(* IEC 61131-3 sources: STEPROBOT/docs/welder_r6_4/source_reference, 3 files *)

(* ---- CommPoll.declaration.original.st ---- *)
(* ================================================================ *)
(* InoProShop 创建方式:                                              *)
(*   右键 Application → 添加对象 → 程序(POU)                        *)
(*   名称: CommPoll, 语言: ST, 类型: PROGRAM                        *)
(*   任务分配: MainTask (1ms周期)                                    *)
(*   说明: 焊机EtherCAT I/O 周期打包/解析                            *)
(*   依赖GVL: GVL_Welder, GVL_CNC                                  *)
(* ================================================================ *)
(*
 * 职责划分:
 *   CNC_Main.st  → 仅设置布尔标志 (g_wWeldOn, g_wRobotReady等)
 *   CommPoll.st  → 每周期: D300拆位→独立BOOL→组装g_byWeldOut
 *                    独立BOOL→组装D308+解析g_byWeldIn
 *
 * 字节映射依据: 奥太EtherCAT通讯协议 2024.7.1
 * PLC数组下标 = 协议字节号 (0-based)
 * ================================================================ *)

PROGRAM CommPoll
VAR
    nTempU16 : UINT;
    nTempI16 : INT;
    byTemp   : BYTE;
    wCtrlPacked : UINT;
    wPrevCtrlPacked : UINT := 16#FFFF;
    bBootInit : BOOL := TRUE;
    rPrevWireAuto : REAL;
    lrPrevWireRun : LREAL;
    bWireParamInit : BOOL := TRUE;
END_VAR

(* ---- CommPoll.implementation.original.st ---- *)
(* Canonical wire parameters: reject NaN/infinity/negative values without
   converting them to integer timer values. No command/enable is generated. *)
IF NOT ((g_rWireStartDelay >= 0.0) AND (g_rWireStartDelay <= 60.0)) THEN
    g_rWireStartDelay := 0.0;
END_IF;
IF NOT ((g_rWireStopDelay >= 0.0) AND (g_rWireStopDelay <= 60.0)) THEN
    g_rWireStopDelay := 0.0;
END_IF;
IF NOT ((g_rWireJogSpeed >= 0.0) AND (g_rWireJogSpeed <= 1000.0)) THEN
    g_rWireJogSpeed := 0.0;
END_IF;
IF NOT ((g_rWireAutoSpeed >= 0.0) AND (g_rWireAutoSpeed <= 1000.0)) THEN
    g_rWireAutoSpeed := 0.0;
END_IF;
IF NOT ((g_fWireFeedSpeed >= 0.0) AND (g_fWireFeedSpeed <= 1000.0)) THEN
    g_fWireFeedSpeed := 0.0;
END_IF;
IF bWireParamInit THEN
    (* Preserve the existing 64-bit setting across restart. *)
    g_rWireAutoSpeed := LREAL_TO_REAL(g_fWireFeedSpeed);
    bWireParamInit := FALSE;
ELSIF g_fWireFeedSpeed <> lrPrevWireRun THEN
    g_rWireAutoSpeed := LREAL_TO_REAL(g_fWireFeedSpeed);
ELSIF g_rWireAutoSpeed <> rPrevWireAuto THEN
    g_fWireFeedSpeed := REAL_TO_LREAL(g_rWireAutoSpeed);
END_IF;
rPrevWireAuto := g_rWireAutoSpeed;
lrPrevWireRun := g_fWireFeedSpeed;
g_dwModbusSignature := 16#4D573031;
g_wModbusMapVersion := 1;
g_dwModbusCycle := g_dwModbusCycle + UDINT#1;
g_wModbusProbeEcho := g_wModbusProbe XOR UINT#16#A55A;

IF bBootInit THEN
    g_wWeldCtrlWord := 0;
    g_wWeldOn := FALSE;
    g_wRobotReady := FALSE;
    g_wGasCheck := FALSE;
    g_bHotWireEnable := FALSE;
    g_bHotWireACMode := FALSE;
    g_bHighFreqDisable := FALSE;
    g_bGunCoolMode := FALSE;
    wPrevCtrlPacked := 0;
    bBootInit := FALSE;
END_IF;

(* ================================================================ *)
(* D300 <-> 独立BOOL 双向合并                                         *)
(* 1. 从独立BOOL打包到临时变量                                        *)
(* 2. 若D300与上次打包值不同(PC写了D300), 则拆位D300→BOOL             *)
(* 3. 再从BOOL打包→D300 (PLC改BOOL也能反映到D300)                     *)
(* ================================================================ *)

wCtrlPacked := 0;
IF g_wWeldOn         THEN wCtrlPacked := wCtrlPacked OR 16#0001; END_IF;
IF g_wRobotReady     THEN wCtrlPacked := wCtrlPacked OR 16#0002; END_IF;
IF g_wGasCheck       THEN wCtrlPacked := wCtrlPacked OR 16#0004; END_IF;
IF g_bHotWireEnable  THEN wCtrlPacked := wCtrlPacked OR 16#0008; END_IF;
IF g_bHotWireACMode  THEN wCtrlPacked := wCtrlPacked OR 16#0010; END_IF;
IF g_bHighFreqDisable THEN wCtrlPacked := wCtrlPacked OR 16#0080; END_IF;
IF g_bGunCoolMode    THEN wCtrlPacked := wCtrlPacked OR 16#0100; END_IF;

IF g_wWeldCtrlWord <> wPrevCtrlPacked THEN
    g_wWeldOn         := (g_wWeldCtrlWord AND 16#0001) <> 0;
    g_wRobotReady     := (g_wWeldCtrlWord AND 16#0002) <> 0;
    g_wGasCheck       := (g_wWeldCtrlWord AND 16#0004) <> 0;
    g_bHotWireEnable  := (g_wWeldCtrlWord AND 16#0008) <> 0;
    g_bHotWireACMode  := (g_wWeldCtrlWord AND 16#0010) <> 0;
    g_bHighFreqDisable := (g_wWeldCtrlWord AND 16#0080) <> 0;
    g_bGunCoolMode    := (g_wWeldCtrlWord AND 16#0100) <> 0;
    wCtrlPacked := g_wWeldCtrlWord;
END_IF;

g_wWeldCtrlWord := wCtrlPacked;
wPrevCtrlPacked := wCtrlPacked;

(* ================================================================ *)
(* 焊机输出 (协议: 焊机的输入数据区, PLC写→焊机读)                    *)
(* g_byWeldOut[0..31] → EtherCAT输出 → 焊机                        *)
(* ================================================================ *)

(* ===== 协议 Byte 0: 控制位 ===== *)
(* bit0(1):  开始焊接 1=起弧 0=停弧                                  *)
(* bit1(2):  机器人准备好 高有效                                      *)
(* bit2(3):  检气 高有效                                              *)
(* bit3-4:   焊机操作模式 00=两步 01=四步 10=反复                     *)
(* bit5-7:   焊机工作模式 000=直流恒流 001=直流脉冲 010=交流恒流       *)
(*           011=交流脉冲 100=直流手弧焊                               *)
byTemp := 0;
IF g_wWeldOn THEN byTemp := byTemp OR 16#01; END_IF;
IF g_wRobotReady THEN byTemp := byTemp OR 16#02; END_IF;
IF g_wGasCheck THEN byTemp := byTemp OR 16#04; END_IF;
nTempU16 := LIMIT(UINT#0, g_wWeldOperMode, UINT#2);
byTemp := byTemp OR SHL(UINT_TO_BYTE(nTempU16), 3);
nTempU16 := LIMIT(UINT#0, g_wWeldWorkMode, UINT#4);
byTemp := byTemp OR SHL(UINT_TO_BYTE(nTempU16), 5);
g_byWeldOut[0] := byTemp;

(* ===== 协议 Byte 1: 辅助控制位 ===== *)
(* bit0(9):  热丝电源使能 1=ON 0=OFF                                  *)
(* bit1(10): 热丝工作模式 0=DC 1=AC                                   *)
(* bit2(11): 备用                                                     *)
(* bit3(12): 点动送丝 (已移除, 送丝通过轴控制) *)
(* bit4(13): 点动抽丝 (已移除, 送丝通过轴控制) *)
(* bit5(14): 备用                                                     *)
(* bit6(15): 高频有无 0=高频 1=提升                                   *)
(* bit7(16): 焊枪模式 0=水冷 1=气冷                                   *)
byTemp := 0;
IF g_bHotWireEnable THEN byTemp := byTemp OR 16#01; END_IF;
IF g_bHotWireACMode THEN byTemp := byTemp OR 16#02; END_IF;
IF g_bHighFreqDisable THEN byTemp := byTemp OR 16#40; END_IF;
IF g_bGunCoolMode THEN byTemp := byTemp OR 16#80; END_IF;
g_byWeldOut[1] := byTemp;

(* ===== 协议 Byte 2: 热丝频率 ===== *)
(* 范围: 20-100 对应20~100Hz (1字节) *)
g_byWeldOut[2] := UINT_TO_BYTE(LIMIT(UINT#20, g_wHotWireFreq, UINT#100));

(* ===== 协议 Byte 3: 热丝电流给定 ===== *)
(* 范围: 0-200 对应0~200A (1字节) *)
g_byWeldOut[3] := UINT_TO_BYTE(LIMIT(UINT#0, g_wHotWireCurrent, UINT#200));

(* ===== 协议 Byte 4-5: 给定电流 (2字节小端, 低字节在前) ===== *)
(* 范围: 40-4000 对应4.0~400.0A *)
nTempU16 := REAL_TO_UINT(LIMIT(4.0, g_wWeldCurrent, 400.0)*10.0);

g_byWeldOut[4] := UINT_TO_BYTE(UINT_TO_USINT(nTempU16 MOD 256));
g_byWeldOut[5] := UINT_TO_BYTE(UINT_TO_USINT(nTempU16 / 256));

(* ===== 协议 Byte 6: 送丝速度 (已移除, 送丝通过轴控制, 写0) ===== *)
g_byWeldOut[6] := 0;

(* ===== 协议 Byte 7: 起弧延迟送丝时间 (已移除, 写0) ===== *)
g_byWeldOut[7] := 0;

(* ===== 协议 Byte 8: 熄弧滞后送丝时间 (已移除, 写0) ===== *)
g_byWeldOut[8] := 0;

(* ===== 协议 Byte 9: 熄弧回抽丝长度 (已移除, 写0) ===== *)
g_byWeldOut[9] := 0;

(* ===== 协议 Byte 10: 点动送丝速度 (已移除, 送丝通过轴控制, 写0) ===== *)
g_byWeldOut[10] := 0;

(* ===== 协议 Byte 11: 通讯异常标志 (控制器填充) ===== *)
g_byWeldOut[11] := g_wCommErrorFlag;

(* ===== 协议 Byte 12: 慢送丝速度 (已移除, 送丝通过轴控制, 写0) ===== *)
g_byWeldOut[12] := 0;

(* ===== 协议 Byte 13-14: 前气时间 (2字节小端, 低字节在前) ===== *)
(* 范围: 1-999 对应0.01~9.99s *)
nTempU16 := REAL_TO_UINT(LIMIT(0.01, g_wFrontGasTime, 9.99)*100.0);
g_byWeldOut[13] := UINT_TO_BYTE(UINT_TO_USINT(nTempU16 MOD 256));
g_byWeldOut[14] := UINT_TO_BYTE(UINT_TO_USINT(nTempU16 / 256));

(* ===== 协议 Byte 15-16: 延气时间 (2字节小端, 低字节在前) ===== *)
(* 范围: 1-600 对应0.1~60.0s *)
nTempU16 := REAL_TO_UINT(LIMIT(0.1, g_wTailGasTime, 60.0)*10.0);
g_byWeldOut[15] := UINT_TO_BYTE(UINT_TO_USINT(nTempU16 MOD 256));
g_byWeldOut[16] := UINT_TO_BYTE(UINT_TO_USINT(nTempU16 / 256));

(* ===== 协议 Byte 17: 爬升时间 ===== *)
(* 范围: 1-100 对应0.1~10.0s (1字节) *)
g_byWeldOut[17] := UINT_TO_BYTE(REAL_TO_UINT(LIMIT(0.1, g_wRampUpTime, 10.0)*10.0));

(* ===== 协议 Byte 18: 衰减时间 ===== *)
(* 范围: 1-150 对应0.1~15.0s (1字节) *)
g_byWeldOut[18] := UINT_TO_BYTE(REAL_TO_UINT(LIMIT(0.1, g_wRampDownTime, 15.0)*10.0));

(* ===== 协议 Byte 19: 脉冲频率 ===== *)
(* 范围: 2-200 对应0.2~20.0Hz (1字节) *)
g_byWeldOut[19] := UINT_TO_BYTE(REAL_TO_UINT(LIMIT(0.2, g_wPulseFreq, 20.0)*10.0));

(* ===== 协议 Byte 20-22: 占空比 + 峰值电流 (交叉编排) ===== *)
(* 占空比: Byte20=低字节, Byte22 bit4-7=高字节低4位 (范围1-999, 12位) *)
(* 峰值电流: Byte21=低字节, Byte22 bit0-3=高字节低4位 (范围50-4000, 12位) *)
(* 占空比 = [Byte22 bit7:4][Byte20] *)
(* 峰值电流 = [Byte22 bit3:0][Byte21] *)
nTempU16 := REAL_TO_UINT(LIMIT(0.1, g_wDutyCycle, 99.9)*10.0);
g_byWeldOut[20] := UINT_TO_BYTE(UINT_TO_USINT(nTempU16 MOD 256));
g_byWeldOut[21] := UINT_TO_BYTE(UINT_TO_USINT(REAL_TO_UINT(LIMIT(5.0, g_wPeakCurrent, 400.0)*10.0) MOD 256));
byTemp := 0;
byTemp := byTemp OR SHL(UINT_TO_BYTE(UINT_TO_USINT(nTempU16 / 256)) AND 16#0F, 4);
byTemp := byTemp OR (UINT_TO_BYTE(UINT_TO_USINT(REAL_TO_UINT(LIMIT(5.0, g_wPeakCurrent, 400.0)*10.0) / 256)) AND 16#0F);
g_byWeldOut[22] := byTemp;

(* ===== 协议 Byte 23-24: 基值电流 (2字节小端, 低字节在前) ===== *)
(* 范围: 50-4000 对应5.0~400.0A *)
nTempU16 := REAL_TO_UINT(LIMIT(5.0, g_wBaseCurrent, 400.0)*10.0);
g_byWeldOut[23] := UINT_TO_BYTE(UINT_TO_USINT(nTempU16 MOD 256));
g_byWeldOut[24] := UINT_TO_BYTE(UINT_TO_USINT(nTempU16 / 256));

(* ===== 协议 Byte 25-26: 起弧电流 (2字节小端, 低字节在前) ===== *)
(* 范围: 50-4000 对应5.0~400.0A *)
nTempU16 := REAL_TO_UINT(LIMIT(5.0, g_wArcStartCurrent, 400.0)*10.0);
g_byWeldOut[25] := UINT_TO_BYTE(UINT_TO_USINT(nTempU16 MOD 256));
g_byWeldOut[26] := UINT_TO_BYTE(UINT_TO_USINT(nTempU16 / 256));

(* ===== 协议 Byte 27-28: 收弧电流 (2字节小端, 低字节在前) ===== *)
(* 范围: 50-4000 对应5.0~400.0A *)
nTempU16 := REAL_TO_UINT(LIMIT(5.0, g_wArcEndCurrent, 400.0)*10.0);
g_byWeldOut[27] := UINT_TO_BYTE(UINT_TO_USINT(nTempU16 MOD 256));
g_byWeldOut[28] := UINT_TO_BYTE(UINT_TO_USINT(nTempU16 / 256));

(* ===== 协议 Byte 29: 交流频率 ===== *)
(* 范围: 40-250 对应40-250Hz (1字节) *)
g_byWeldOut[29] := UINT_TO_BYTE(LIMIT(UINT#40, g_wACFreq, UINT#250));

(* ===== 协议 Byte 30: 清理比例 ===== *)
(* 范围: 90-180 对应40~-50 (1字节) *)
nTempI16 := 130 - UINT_TO_INT(LIMIT(UINT#90, g_wCleanRatio, UINT#180));
g_byWeldOut[30] := INT_TO_BYTE(nTempI16);

(* ===== 协议 Byte 31: 交流偏置 ===== *)
(* 范围: 90-180 对应40~-50 (1字节) *)
nTempI16 := 130 - UINT_TO_INT(LIMIT(UINT#90, g_wACBias, UINT#180));
g_byWeldOut[31] := INT_TO_BYTE(nTempI16);

(* ================================================================ *)
(* 焊机输入 (协议: 焊机输出数据区, 焊机写→PLC读)                      *)
(* g_byWeldIn[0..31] ← EtherCAT输入 ← 焊机                          *)
(* ================================================================ *)

(* ===== 协议输入 Byte 0: 状态位 ===== *)
(* bit0: 引弧成功 高有效                                              *)
(* bit1: 焊机准备好 高有效                                            *)
(* bit2: 预留                                                         *)
(* bit3: 电流有无 高有效                                              *)
(* EtherCAT 输入映射别名 → 协议数组。保持原有 Byte 0..31 定义。 *)
g_byWeldIn[0] := g_byWeldInMap01;
g_byWeldIn[1] := g_byWeldInMap02;
g_byWeldIn[2] := g_byWeldInMap03;
g_byWeldIn[3] := g_byWeldInMap04;
g_byWeldIn[4] := g_byWeldInMap05;
g_byWeldIn[5] := g_byWeldInMap06;
g_byWeldIn[6] := g_byWeldInMap07;
g_byWeldIn[7] := g_byWeldInMap08;
g_byWeldIn[8] := g_byWeldInMap09;
g_byWeldIn[9] := g_byWeldInMap10;
g_byWeldIn[10] := g_byWeldInMap11;
g_byWeldIn[11] := g_byWeldInMap12;
g_byWeldIn[12] := g_byWeldInMap13;
g_byWeldIn[13] := g_byWeldInMap14;
g_byWeldIn[14] := g_byWeldInMap15;
g_byWeldIn[15] := g_byWeldInMap16;
g_byWeldIn[16] := g_byWeldInMap17;
g_byWeldIn[17] := g_byWeldInMap18;
g_byWeldIn[18] := g_byWeldInMap19;
g_byWeldIn[19] := g_byWeldInMap20;
g_byWeldIn[20] := g_byWeldInMap21;
g_byWeldIn[21] := g_byWeldInMap22;
g_byWeldIn[22] := g_byWeldInMap23;
g_byWeldIn[23] := g_byWeldInMap24;
g_byWeldIn[24] := g_byWeldInMap25;
g_byWeldIn[25] := g_byWeldInMap26;
g_byWeldIn[26] := g_byWeldInMap27;
g_byWeldIn[27] := g_byWeldInMap28;
g_byWeldIn[28] := g_byWeldInMap29;
g_byWeldIn[29] := g_byWeldInMap30;
g_byWeldIn[30] := g_byWeldInMap31;
g_byWeldIn[31] := g_byWeldInMap32;

g_bWeldArcOK      := (g_byWeldIn[0] AND 16#01) <> 0;
g_bWeldReady      := (g_byWeldIn[0] AND 16#02) <> 0;
g_bWeldHasCurrent     := (g_byWeldIn[0] AND 16#08) <> 0;

(* ===== 协议输入 Byte 1: 报警位 ===== *)
(* bit0: 预留                                                         *)
(* bit1: 焊枪开关异常 高有效                                          *)
(* bit2: 焊机热保护 高有效                                            *)
(* bit3: 缺水保护 高有效                                              *)
(* bit4: 热丝电源热保护 高有效                                        *)
(* bit5: 热丝电源通讯保护 高有效 (控制器填充)                          *)
g_bGunSwitchFault    := (g_byWeldIn[1] AND 16#02) <> 0;
g_bWeldThermalProtect := (g_byWeldIn[1] AND 16#04) <> 0;
g_bWaterProtect   := (g_byWeldIn[1] AND 16#08) <> 0;
g_bWirePSThermal  := (g_byWeldIn[1] AND 16#10) <> 0;
g_bWirePSCommFault:= (g_byWeldIn[1] AND 16#20) <> 0;

(* ===== 报警组合 ===== *)
g_bWeldFault := g_bWeldThermalProtect
              OR g_bGunSwitchFault
              OR g_bWaterProtect
              OR g_bWirePSThermal
              OR g_bWirePSCommFault;

IF g_bWeldFault THEN
    g_rWeldFaultCode := BYTE_TO_UINT(g_byWeldIn[1]);
ELSE
    g_rWeldFaultCode := 0;
END_IF;

IF NOT g_bWeldReady OR g_bWeldFault THEN
    g_wWeldOn := FALSE;
    g_wWeldCtrlWord := g_wWeldCtrlWord AND 16#FFFE;
    wPrevCtrlPacked := wPrevCtrlPacked AND 16#FFFE;
    g_byWeldOut[0] := g_byWeldOut[0] AND 16#FE;
END_IF;

(* ===== EtherCAT 输出映射别名同步 ===== *)
(* 放在未就绪/故障联锁之后，确保停弧命令在本周期立即写入PDO。 *)
g_byWeldOutMap01 := g_byWeldOut[0];
g_byWeldOutMap02 := g_byWeldOut[1];
g_byWeldOutMap03 := g_byWeldOut[2];
g_byWeldOutMap04 := g_byWeldOut[3];
g_byWeldOutMap05 := g_byWeldOut[4];
g_byWeldOutMap06 := g_byWeldOut[5];
g_byWeldOutMap07 := g_byWeldOut[6];
g_byWeldOutMap08 := g_byWeldOut[7];
g_byWeldOutMap09 := g_byWeldOut[8];
g_byWeldOutMap10 := g_byWeldOut[9];
g_byWeldOutMap11 := g_byWeldOut[10];
g_byWeldOutMap12 := g_byWeldOut[11];
g_byWeldOutMap13 := g_byWeldOut[12];
g_byWeldOutMap14 := g_byWeldOut[13];
g_byWeldOutMap15 := g_byWeldOut[14];
g_byWeldOutMap16 := g_byWeldOut[15];
g_byWeldOutMap17 := g_byWeldOut[16];
g_byWeldOutMap18 := g_byWeldOut[17];
g_byWeldOutMap19 := g_byWeldOut[18];
g_byWeldOutMap20 := g_byWeldOut[19];
g_byWeldOutMap21 := g_byWeldOut[20];
g_byWeldOutMap22 := g_byWeldOut[21];
g_byWeldOutMap23 := g_byWeldOut[22];
g_byWeldOutMap24 := g_byWeldOut[23];
g_byWeldOutMap25 := g_byWeldOut[24];
g_byWeldOutMap26 := g_byWeldOut[25];
g_byWeldOutMap27 := g_byWeldOut[26];
g_byWeldOutMap28 := g_byWeldOut[27];
g_byWeldOutMap29 := g_byWeldOut[28];
g_byWeldOutMap30 := g_byWeldOut[29];
g_byWeldOutMap31 := g_byWeldOut[30];
g_byWeldOutMap32 := g_byWeldOut[31];

(* ===== 协议输入 Byte 4-5: 实际焊接电压 (2字节小端, 0.1V分辨率) ===== *)
(* 范围: 0-1000 对应0~100.0V *)
nTempU16 := BYTE_TO_UINT(g_byWeldIn[4]) + BYTE_TO_UINT(g_byWeldIn[5]) * 256;
g_rWeldVoltageAct := UINT_TO_REAL(nTempU16) * 0.1;

(* ===== 协议输入 Byte 6-7: 实际焊接电流 (2字节小端, 0.1A分辨率) ===== *)
(* 范围: 0~400 对应0~400A *)
nTempU16 := BYTE_TO_UINT(g_byWeldIn[6]) + BYTE_TO_UINT(g_byWeldIn[7]) * 256;
g_rWeldCurrentAct := UINT_TO_REAL(nTempU16) * 0.1;

(* ===== 协议输入 Byte 8-9: 实际热丝焊接电流 (2字节小端, 10A分辨率) ===== *)
(* 范围: 0~20 对应0~200A *)
nTempU16 := BYTE_TO_UINT(g_byWeldIn[8]) + BYTE_TO_UINT(g_byWeldIn[9]) * 256;
g_rHotWireCurrentAct := UINT_TO_REAL(nTempU16) * 10.0;

(* ===== 协议输入 Byte 10-11: 送丝速度反馈 (已移除, 送丝通过轴控制) ===== *)

(* ===== 组装输入状态字 (PC通过D500读取) ===== *)
g_wWeldInStatus := 0;
IF g_bWeldArcOK      THEN g_wWeldInStatus := g_wWeldInStatus OR 16#0001; END_IF;
IF g_bWeldReady      THEN g_wWeldInStatus := g_wWeldInStatus OR 16#0002; END_IF;
IF g_bGunSwitchFault THEN g_wWeldInStatus := g_wWeldInStatus OR 16#0004; END_IF;
IF g_bWeldThermalProtect THEN g_wWeldInStatus := g_wWeldInStatus OR 16#0008; END_IF;
IF g_bWaterProtect   THEN g_wWeldInStatus := g_wWeldInStatus OR 16#0010; END_IF;
IF g_bWirePSThermal  THEN g_wWeldInStatus := g_wWeldInStatus OR 16#0020; END_IF;
IF g_bWirePSCommFault THEN g_wWeldInStatus := g_wWeldInStatus OR 16#0040; END_IF;
IF g_bWeldFault      THEN g_wWeldInStatus := g_wWeldInStatus OR 16#0080; END_IF;
IF g_bWeldHasCurrent     THEN g_wWeldInStatus := g_wWeldInStatus OR 16#0100; END_IF;

(* ================================================================ *)
(* D308 独立BOOL → 打包字 (PLC内部 → PC读D308)                         *)
(* CommPoll每周期从独立BOOL组装到g_wWeldStatusWord供PC读取             *)
(* ================================================================ *)
g_wWeldStatusWord := 0;
IF g_bWeldArcOK      THEN g_wWeldStatusWord := g_wWeldStatusWord OR 16#0001; END_IF;
IF g_bWeldReady      THEN g_wWeldStatusWord := g_wWeldStatusWord OR 16#0002; END_IF;
IF g_bWeldHasCurrent     THEN g_wWeldStatusWord := g_wWeldStatusWord OR 16#0004; END_IF;
IF g_bGunSwitchFault THEN g_wWeldStatusWord := g_wWeldStatusWord OR 16#0008; END_IF;
IF g_bWeldThermalProtect THEN g_wWeldStatusWord := g_wWeldStatusWord OR 16#0010; END_IF;
IF g_bWaterProtect   THEN g_wWeldStatusWord := g_wWeldStatusWord OR 16#0020; END_IF;
IF g_bWirePSThermal  THEN g_wWeldStatusWord := g_wWeldStatusWord OR 16#0040; END_IF;
IF g_bWirePSCommFault THEN g_wWeldStatusWord := g_wWeldStatusWord OR 16#0080; END_IF;
IF g_bWeldFault      THEN g_wWeldStatusWord := g_wWeldStatusWord OR 16#0100; END_IF;

(* ================================================================ *)
(* 激光距离读取和转换                                                *)
(* 从%IW50读取激光距离原始INT值, 转换为实际距离并存入寄存器            *)
(* 转换公式: 实际距离 = 原始值 / 100 + 50                             *)
(* D522 = g_rLaserDistance (REAL, PC可通过Modbus读取)                   *)
(* ================================================================ *)
g_rLaserDistance := INT_TO_REAL(g_iLaserDistanceRaw) / 100.0 + 50.0;

(* ---- GVL_Welders.original.st ---- *)
(* EtherCAT -9 welder: 32-byte RxPDO/TxPDO use symbolic channel mappings; no fixed IEC addresses. *)
(* ================================================================ *)
(* InoProShop 创建方式:                                              *)
(*   右键 Application → 添加对象 → 全局变量表(GVL)                    *)
(*   名称: GVL_Welders                                               *)
(*   说明: 奥太焊机 EtherCAT 通讯接口全局变量                         *)
(*   依赖: 无                                                        *)
(*   修订: 布尔变量使用独立%MW地址 (D300控制=%MW101~109)               *)
(*         (D308状态=%MW111~119), InoProShop不支持BOOL位打包         *)
(*         新增 %MW300/%MW308 作为Modbus从站打包字映射 (方案C)         *)
(* ================================================================ *)
(*
 * EtherCAT通讯协议 (奥太 2024.7.1)
 *
 * EtherCAT输出 (PLC→焊机): g_byWeldOut[0..31] → 地址-9焊机RxPDO (32字节)
 *   协议字节0~31 = PLC数组下标0~31 (一一对应)
 *
 * EtherCAT输入 (焊机→PLC): g_byWeldIn[0..31] ← 地址-9焊机TxPDO (32字节)
 *   协议字节0~31 = PLC数组下标0~31 (一一对应)
 *
 * 数据流:
 *   PC(Modbus写D300) → g_wWeldCtrlWord (打包字)
 *       → CommPoll.st拆位 → g_wWeldOn等独立BOOL
 *       → CommPoll.st组装 → g_byWeldOut → EtherCAT → 焊机
 *   焊机 → EtherCAT → g_byWeldIn
 *       → CommPoll.st解析 → g_bWeldArcOK等独立BOOL
 *       → CommPoll.st组装 → g_wWeldStatusWord → PC(Modbus读D308)
 *
 * Modbus寄存器布局:
 *   D300 (%MW300): 焊机控制输出标志位 (16位打包字, CommPoll双向映射)
 *     独立BOOL: g_wWeldOn(%MW101) ~ g_bGunCoolMode(%MW109)
 *   D302      : 焊机操作模式 (UINT)
 *   D304      : 焊机工作模式 (UINT)
 *   D306      : 通讯异常标志 (BYTE, 控制器填充)
 *   D308 (%MW308): 焊机输入状态标志位 (16位打包字, CommPoll组装)
 *     独立BOOL: g_bWeldArcOK(%MW111) ~ g_bWeldFault(%MW119)
 *   D400-D444 : 焊接参数 (各参数见注释)
 *   D500      : 焊机输入状态字 (16位打包, CommPoll从独立BOOL组装)
 *   D502-D518 : 焊机输入反馈值
 *
 * 注意: Modbus从站配置需包含 D300-D306 和 D308 映射范围
 *       D300=%MW300, D308=%MW308 均为打包字, PC按位操作
 * ================================================================ *)

(* ================================================================= *)
(* 焊机控制输出标志位 → 协议 Byte 0 / Byte 1 位域                     *)
(* Modbus: D300 (%MW300, 16位), bit0~8 对应9个布尔量                  *)
(* ================================================================= *)

(*
 * 协议 Byte 0 位域:
 *   bit0(1):  开始焊接       1=起弧 0=停弧 [危险, 高有效]
 *   bit1(2):  机器人准备好   上位机接收到焊机数据, 通讯正常, 高有效
 *   bit2(3):  检气           高有效
 *   bit3-4:   焊机操作模式   00=两步 01=四步 10=反复
 *   bit5-7:   焊机工作模式   000=直流恒流 001=直流脉冲 010=交流恒流
 *             011=交流脉冲 100=直流手弧焊
 *
 * 协议 Byte 1 位域:
 *   bit0(9):  热丝电源使能   1=ON 0=OFF
 *   bit1(10): 热丝工作模式   0=DC 1=AC
 *   bit2(11): 备用
 *   bit3(12): 点动送丝       高有效, 丝检时使用, 电平信号
 *   bit4(13): 点动抽丝       高有效, 丝检时使用, 电平信号
 *   bit5(14): 备用
 *   bit6(15): 高频有无       0=高频 1=提升
 *   bit7(16): 焊枪模式       0=水冷 1=气冷
 *)

(* --- 协议 Byte 11: 通讯异常标志 (控制器填充) --- *)
(*
 * 协议 Byte 11 位域:
 *   bit0(89):  机器人→CAN控制器通信异常 (控制器填充, 焊机显示E84)
 *             注: 500ms内无机器人准备好信号将触发此异常
 *   bit1-3:    预留
 *   bit4(93):  焊机→CAN控制器通信异常 (控制器填充, 焊机显示E85)
 *   bit5-7:    预留
 *)

(* ================================================================= *)
(* 焊接参数 Modbus 接收 (D400~D444)                                  *)
(* PC写入Modbus寄存器 → CommPoll.st读取并组装到g_byWeldOut             *)
//

(* --- 协议 Byte 20-22: 占空比 + 峰值电流 (交叉编排) --- *)
(*
 * 占空比: Byte20=低字节, Byte22 bit4-7=高4位 (12位)
 * 峰值电流: Byte21=低字节, Byte22 bit0-3=高4位 (12位)
 * g_wDutyCycle为REAL, 存实际百分比(如50.0=50.0%, 3.5=3.5%)
 * CommPoll内部 ×10 → 协议值1~999 → 0.1%~99.9%
 * 峰值电流 = [Byte22 bit3:0][Byte21]   范围50~4000 → 5.0~400.0A
 *)

 (* ================================================================= *)
(* 焊机输入状态标志位 → 协议输入 Byte 0 / Byte 1 位域                  *)
(* Modbus: D308 (%MW308, 16位), bit0~8 对应9个布尔量                  *)
(* 由 CommPoll.st 每周期从 g_byWeldIn 解析写入                        *)
(* ================================================================= *)
(*
 * 协议输入 Byte 0:
 *   bit0: 引弧成功     高有效
 *   bit1: 焊机准备好   高有效
 *   bit2: 预留
 *   bit3: 电流有无     高有效
 *   bit4-7: 预留
 *
 * 协议输入 Byte 1:
 *   bit0: 预留
 *   bit1: 焊枪开关异常   高有效
 *   bit2: 焊机热保护     高有效
 *   bit3: 缺水保护       高有效
 *   bit4: 热丝电源热保护 高有效
 *   bit5: 热丝电源通讯保护 高有效 (控制器填充)
 *   bit6-7: 预留
 * ================================================================= *)

 (* ================================================================= *)
(* 输入状态字 (打包, PC通过Modbus D500读取)                            *)
(* 由 CommPoll.st 每周期从各布尔标志位组装写入                          *)
(* ================================================================= *)
(*
 * g_wWeldInStatus 位域 (CommPoll从独立BOOL组装):
 *   bit0:  引弧成功         (g_bWeldArcOK)
 *   bit1:  焊机准备好       (g_bWeldReady)
 *   bit2:  焊枪开关异常     (g_bGunSwitchFault)
 *   bit3:  焊机热保护       (g_bWeldThermalProtect)
 *   bit4:  缺水保护         (g_bWaterProtect)
 *   bit5:  热丝电源热保护   (g_bWirePSThermal)
 *   bit6:  热丝电源通讯保护 (g_bWirePSCommFault)
 *   bit7:  总报警           (g_bWeldFault)
 *   bit8:  电流有无         (g_bWeldHasCurrent)
 *)

(* ================================================================= *)
(* 输入反馈值 (PC通过Modbus读取)                                       *)
(* 由 CommPoll.st 每周期从 g_byWeldIn 解析写入                        *)
(* ================================================================= *)
VAR_GLOBAL
    (* EtherCAT输出 → 焊机输入数据区 (32字节) *)
    g_byWeldOut : ARRAY[0..31] OF BYTE;
    (* EtherCAT输入 ← 焊机输出数据区 (32字节) *)
    g_byWeldIn : ARRAY[0..31] OF BYTE;

    (*
     * EtherCAT 映射别名。
     * InoProShop 的 I/O 映射器要求变量是单一标识符，不接受数组下标；
     * CommPoll 在这些别名与协议数组之间逐周期同步，协议字节编号保持不变。
     *)
    g_byWeldOutMap01 : BYTE;
    g_byWeldOutMap02 : BYTE;
    g_byWeldOutMap03 : BYTE;
    g_byWeldOutMap04 : BYTE;
    g_byWeldOutMap05 : BYTE;
    g_byWeldOutMap06 : BYTE;
    g_byWeldOutMap07 : BYTE;
    g_byWeldOutMap08 : BYTE;
    g_byWeldOutMap09 : BYTE;
    g_byWeldOutMap10 : BYTE;
    g_byWeldOutMap11 : BYTE;
    g_byWeldOutMap12 : BYTE;
    g_byWeldOutMap13 : BYTE;
    g_byWeldOutMap14 : BYTE;
    g_byWeldOutMap15 : BYTE;
    g_byWeldOutMap16 : BYTE;
    g_byWeldOutMap17 : BYTE;
    g_byWeldOutMap18 : BYTE;
    g_byWeldOutMap19 : BYTE;
    g_byWeldOutMap20 : BYTE;
    g_byWeldOutMap21 : BYTE;
    g_byWeldOutMap22 : BYTE;
    g_byWeldOutMap23 : BYTE;
    g_byWeldOutMap24 : BYTE;
    g_byWeldOutMap25 : BYTE;
    g_byWeldOutMap26 : BYTE;
    g_byWeldOutMap27 : BYTE;
    g_byWeldOutMap28 : BYTE;
    g_byWeldOutMap29 : BYTE;
    g_byWeldOutMap30 : BYTE;
    g_byWeldOutMap31 : BYTE;
    g_byWeldOutMap32 : BYTE;

    g_byWeldInMap01 : BYTE;
    g_byWeldInMap02 : BYTE;
    g_byWeldInMap03 : BYTE;
    g_byWeldInMap04 : BYTE;
    g_byWeldInMap05 : BYTE;
    g_byWeldInMap06 : BYTE;
    g_byWeldInMap07 : BYTE;
    g_byWeldInMap08 : BYTE;
    g_byWeldInMap09 : BYTE;
    g_byWeldInMap10 : BYTE;
    g_byWeldInMap11 : BYTE;
    g_byWeldInMap12 : BYTE;
    g_byWeldInMap13 : BYTE;
    g_byWeldInMap14 : BYTE;
    g_byWeldInMap15 : BYTE;
    g_byWeldInMap16 : BYTE;
    g_byWeldInMap17 : BYTE;
    g_byWeldInMap18 : BYTE;
    g_byWeldInMap19 : BYTE;
    g_byWeldInMap20 : BYTE;
    g_byWeldInMap21 : BYTE;
    g_byWeldInMap22 : BYTE;
    g_byWeldInMap23 : BYTE;
    g_byWeldInMap24 : BYTE;
    g_byWeldInMap25 : BYTE;
    g_byWeldInMap26 : BYTE;
    g_byWeldInMap27 : BYTE;
    g_byWeldInMap28 : BYTE;
    g_byWeldInMap29 : BYTE;
    g_byWeldInMap30 : BYTE;
    g_byWeldInMap31 : BYTE;
    g_byWeldInMap32 : BYTE;

	(* D520 | 激光距离 (原始INT值, 从%IW50读取) *)
	(* --- 激光距离原始值 --- *)
	g_iLaserDistanceRaw : INT;
END_VAR

VAR_GLOBAL RETAIN PERSISTENT

(* D300 | 控制标志位打包字 (PC通过Modbus读写, CommPoll每周期双向映射) *)
g_wWeldCtrlWord    AT %MW300 : UINT := 0;

(* D300 bit0 | 独立BOOL | 开始焊接 1=起弧 0=停弧 [危险, 高有效] *)
g_wWeldOn AT %MW101 : BOOL := FALSE;

(* D300 bit1 | 独立BOOL | 机器人准备好, 高有效 *)
g_wRobotReady AT %MW102 : BOOL := FALSE;
(* D300 bit2 | 独立BOOL | 检气, 高有效 *)
g_wGasCheck AT %MW103 : BOOL := FALSE;

(* D300 bit3 | 独立BOOL | 热丝电源使能 1=ON 0=OFF *)
g_bHotWireEnable AT %MW104 : BOOL := FALSE;

(* D300 bit4 | 独立BOOL | 热丝工作模式 0=DC 1=AC *)
g_bHotWireACMode AT %MW105 : BOOL := FALSE;

(* D300 bit7 | 独立BOOL | 高频有无 0=高频 1=提升 *)
g_bHighFreqDisable AT %MW108 : BOOL := FALSE;

(* D300 bit8 | 独立BOOL | 焊枪模式 0=水冷 1=气冷 *)
g_bGunCoolMode AT %MW109 : BOOL := FALSE;

(* D302 | 协议Byte0 bit3-4 | 焊机操作模式 0=两步 1=四步 2=反复 *)
g_wWeldOperMode    AT %MW302 : UINT := 0;

(* D304 | 协议Byte0 bit5-7 | 焊机工作模式 0=直流恒流 1=直流脉冲 2=交流恒流 *)
(*                           3=交流脉冲 4=直流手弧焊 *)
g_wWeldWorkMode    AT %MW304 : UINT := 1;

(* D306 | 协议Byte11 | 通讯异常标志, 控制器填充, 默认0 *)
g_wCommErrorFlag   AT %MW306 : BYTE;

(* D414 | 协议Byte2 bit0-7 | 热丝频率, 范围20~100, 对应20~100Hz (直通) *)
g_wHotWireFreq     AT %MW414 : UINT := 50;

(* D416 | 协议Byte3 bit0-7 | 热丝电流给定, 范围0~200, 对应0~200A (直通) *)
g_wHotWireCurrent  AT %MW416 : UINT := 150;

(* D400 | 协议Byte4-5 | 给定电流, 实际A, 例: 100.0表示100.0A *)
(* CommPoll内部 ×10 → 协议值(范围40~4000, 对应4.0~400.0A), 占D400-D401 *)
g_wWeldCurrent     AT %MW400 : REAL := 100.0;

(* Local wire-feed axis parameters. Speeds are mm/s; delays are seconds.
   D412 and D1202 set the same automatic speed; a changed D1202 has priority.
   D410 > 0 overrides D2104 for axis 4 jog; zero uses D2104 for compatibility. *)
g_rWireStartDelay  AT %MW404 : REAL := 0.0;
g_rWireStopDelay   AT %MW406 : REAL := 0.0;
g_rWireJogSpeed    AT %MW410 : REAL := 0.0;
g_rWireAutoSpeed   AT %MW412 : REAL := 0.0;

(* D420 | 协议Byte13-14 | 前气时间, 实际s, 例: 5.0表示5.00s *)
(* CommPoll内部 ×100 → 协议值(范围1~999, 对应0.01~9.99s), 占D420-D421 *)
g_wFrontGasTime    AT %MW420 : REAL := 0.01;

(* D422 | 协议Byte15-16 | 延气时间, 实际s, 例: 3.0表示3.0s *)
(* CommPoll内部 ×10 → 协议值(范围1~600, 对应0.1~60.0s), 占D422-D423 *)
g_wTailGasTime     AT %MW422 : REAL := 0.2;

(* D424 | 协议Byte17 bit0-7 | 爬升时间, 实际s, 例: 5.0表示5.0s *)
(* CommPoll内部 ×10 → 协议值(范围1~100, 对应0.1~10.0s), 占D424-D425 *)
g_wRampUpTime      AT %MW424 : REAL := 0.5;

(* D426 | 协议Byte18 bit0-7 | 衰减时间, 实际s, 例: 5.0表示5.0s *)
(* CommPoll内部 ×10 → 协议值(范围1~150, 对应0.1~15.0s) *)
g_wRampDownTime    AT %MW426 : REAL := 0.2;

(* D428 | 协议Byte19 bit0-7 | 脉冲频率, 实际Hz, 例: 5.0表示5.0Hz *)
(* CommPoll内部 ×10 → 协议值(范围2~200, 对应0.2~20.0Hz), 占D428-D429 *)
g_wPulseFreq       AT %MW428 : REAL := 0.5;

(* D430 | 协议Byte20+22 bit4-7 | 占空比, 实际百分比, 例: 50.0表示50.0% *)
(* CommPoll内部 ×10 → 协议值(范围1~999, 对应0.1%~99.9%), 占D430-D431 *)
g_wDutyCycle       AT %MW430 : REAL := 50.0;

(* D432 | 协议Byte21+22 bit0-3 | 峰值电流, 实际A, 例: 150.0表示150.0A *)
(* CommPoll内部 ×10 → 协议值(范围50~4000, 对应5.0~400.0A), 占D432-D433 *)
g_wPeakCurrent     AT %MW432 : REAL := 100.0;

(* D434 | 协议Byte23-24 | 基值电流, 实际A, 例: 30.0表示30.0A *)
(* CommPoll内部 ×10 → 协议值(范围50~4000, 对应5.0~400.0A), 占D434-D435 *)
g_wBaseCurrent     AT %MW434 : REAL := 30.0;

(* D436 | 协议Byte25-26 | 起弧电流, 实际A, 例: 100.0表示100.0A *)
(* CommPoll内部 ×10 → 协议值(范围50~4000, 对应5.0~400.0A), 占D436-D437 *)
(* --- 协议 Byte 25-26: 起弧电流 (2字节小端, 低字节在前) --- *)
g_wArcStartCurrent AT %MW436 : REAL;

(* D438 | 协议Byte27-28 | 收弧电流, 实际A, 例: 100.0表示100.0A *)
(* CommPoll内部 ×10 → 协议值(范围50~4000, 对应5.0~400.0A), 占D438-D439 *)
(* --- 协议 Byte 27-28: 收弧电流 (2字节小端, 低字节在前) --- *)
g_wArcEndCurrent   AT %MW438 : REAL;

(* D440 | 协议Byte29 bit0-7 | 交流频率, 范围40~250, 对应40~250Hz (直通) *)
(* --- 协议 Byte 29: 交流频率 --- *)
g_wACFreq          AT %MW440 : UINT;

(* D442 | 协议Byte30 bit0-7 | 清理比例, 范围90~180, 对应40~-50 *)
(* 协议转换: Byte30 = -1 × D442 + 130 *)
(* 例: D442=90 → Byte30=40, D442=130 → Byte30=0, D442=180 → Byte30=-50 *)
(* --- 协议 Byte 30: 清理比例 --- *)
g_wCleanRatio      AT %MW442 : UINT;

(* D444 | 协议Byte31 bit0-7 | 交流偏置, 范围90~180, 对应40~-50 *)
(* 协议转换: Byte31 = -1 × D444 + 130 *)
(* 例: D444=90 → Byte31=40, D444=130 → Byte31=0, D444=180 → Byte31=-50 *)
(* --- 协议 Byte 31: 交流偏置 --- *)
g_wACBias          AT %MW444 : UINT;

(* D308 | 输入状态打包字 (PC通过Modbus读取, CommPoll每周期从独立BOOL组装) *)
g_wWeldStatusWord  AT %MW308 : UINT;

(* D308 bit0 | 独立BOOL | 引弧成功, 高有效 *)
g_bWeldArcOK AT %MW111 : BOOL;

(* D308 bit1 | 独立BOOL | 焊机准备好, 高有效 *)
g_bWeldReady AT %MW112 : BOOL;

(* D308 bit2 | 独立BOOL | 电流有无, 高有效 *)
g_bWeldHasCurrent AT %MW113 : BOOL;

(* D308 bit3 | 独立BOOL | 焊枪开关异常, 高有效 *)
g_bGunSwitchFault AT %MW114 : BOOL;

(* D308 bit4 | 独立BOOL | 焊机热保护, 高有效 *)
g_bWeldThermalProtect AT %MW115 : BOOL;

(* D308 bit5 | 独立BOOL | 缺水保护, 高有效 *)
g_bWaterProtect AT %MW116 : BOOL;

(* D308 bit6 | 独立BOOL | 热丝电源热保护, 高有效 *)
g_bWirePSThermal AT %MW117 : BOOL;

(* D308 bit7 | 独立BOOL | 热丝电源通讯保护, 高有效, 控制器填充 *)
g_bWirePSCommFault AT %MW118 : BOOL;

(* D308 bit8 | 独立BOOL | 组合报警, 包含焊枪开关/热保护/缺水/热丝电源故障 *)
g_bWeldFault AT %MW119 : BOOL;

(* D500 | 焊机输入状态字 (16位打包, 详见位域定义) *)
g_wWeldInStatus    AT %MW500 : UINT;

(* D502-D503 | 协议输入Byte4-5 | 实际焊接电压, 0.1V分辨率 *)
(* --- 协议输入 Byte 4-5: 实际焊接电压 (2字节小端, 0.1V分辨率) --- *)
(* 范围: 0~1000 → 0~100.0V *)
g_rWeldVoltageAct    AT %MW502 : REAL;

(* D506-D507 | 协议输入Byte6-7 | 实际焊接电流, 0.1A分辨率 *)
(* --- 协议输入 Byte 6-7: 实际焊接电流 (2字节小端, 0.1A分辨率) --- *)
(* 范围: 0~400 → 0~400A *)
g_rWeldCurrentAct    AT %MW506 : REAL;

(* D510-D511 | 协议输入Byte8-9 | 实际热丝焊接电流, 10A分辨率 *)
(* --- 协议输入 Byte 8-9: 实际热丝焊接电流 (2字节小端, 10A分辨率) --- *)
(* 范围: 0~20 → 0~200A *)
g_rHotWireCurrentAct AT %MW510 : REAL;

(* D518 | 协议输入Byte1原始值 | 报警码, 报警时记录协议输入Byte1原始值 *)
(* --- 报警原始字节 --- *)
g_rWeldFaultCode     AT %MW518 : UINT;

(* D522 | 激光距离 (实际距离mm, 原始值/100+50) *)
(* --- 激光距离实际值 --- *)
g_rLaserDistance AT %MW522 : REAL := 50.0;

(* ================================================================= *)
(* 协议输入预留字节 (协议保留, 当前未使用)                               *)
(*   协议输入 Byte 2-3: 预留                                          *)
(*   协议输入 Byte 12:  预留                                          *)
(* ================================================================= *)

END_VAR
